(* IEC 61131-3 sources: Elmo_Master/Lasal_PRG/Welcon8Axis_EtherCAT_Test_With_RobotAxis/Class/SafetyCDIAS_Base (part 6) *)

  //Check pointer
  if pData then
    //Length of Firmwareversion (HDINT) -> 8Byte +1 byte zero termination
    if Length >= 9 then
      _itoa(udNumber:=FW_Version, pString:=pData);
    else
      pData^ := 0;
    end_if;
  end_if;

END_FUNCTION

FUNCTION VIRTUAL GLOBAL SafetyCDIAS_Base::GetDiagConnect::NewInst
	VAR_INPUT
		pPara 	  : ^CmdStruct;
		pResult 	: ^Results;
	END_VAR
	VAR_OUTPUT
		ret_code 	: IprStates;
	END_VAR

	ret_code := READY;

	CASE pPara^.uiCmd OF

    CMD_SM_DIAG_GET_INFO:

      //Subcommand
      case pPara^.aPara[0] of
//*****************************************************************************
        SBCMD_SM_DIAG_GET_INFO:
          pResult^.aData[0] :=  GetDiagInfo(pDiagInfo:=(pPara^.aPara[1])$^SafetyDiagInfo);

//*****************************************************************************
        SBCMD_SM_DIAG_GET_STATE:
          pResult^.aData[0] :=  GetDiagState(pDiagState:=(pPara^.aPara[1])$^SafetyDiagState);

//*****************************************************************************
        SBCMD_SM_DIAG_FETCH_INFO:
          //Fetch Diag Info for uCx
          FetchDiagInfo(ucChoice:=pPara^.aPara[1]$USINT);

//*****************************************************************************
        SBCMD_SM_DIAG_FETCH_STATE:
          FetchDiagState();

//*****************************************************************************
        SBCMD_SM_DIAG_IS_SAVE_LOG_ACTIVE:
          pResult^.aData[0] := SaveLogActive();

//*****************************************************************************
        SBCMD_SM_DIAG_SAVE_LOGFILE:
          pResult^.aData[0] := (SaveLog(ucChoice:=(pPara^.aPara[1])$USINT, pDPNE:=(pPara^.aPara[2])$^CHAR))$USINT;

//*****************************************************************************
        SBCMD_SM_DIAG_GET_SAVE_LOGFILE_STATE:
          pResult^.aData[0] := DiagVars.SavingLogSuccessful$USINT;

//*****************************************************************************
        SBCMD_SM_DIAG_GET_SAFETY_NUMBER:
          pResult^.aData[0]$UDINT := SafetyNumber;

//*****************************************************************************
        SBCMD_SM_DIAG_GET_SAFETY_STATE:
          pResult^.aData[0] := ClassState$USINT;

//*****************************************************************************
        SBCMD_SM_DIAG_IS_DIAGNOSE_AVAILABLE:
          pResult^.aData[0] := TRUE;

//*****************************************************************************
        SBCMD_SM_DIAG_GET_CHANNEL_INFO:
          pResult^.aData[0] := GetChannelInfo(pErrorMemUser:=(pPara^.aPara[1])$^UINT, pErrorMem:=#aErrorMem[1], ErrorDataLength:=aErrorMem[0] - 1);
          pResult^.aData[1] := aErrorMem[0] - 1;

//*****************************************************************************
        SBCMD_SM_DIAG_FETCH_CHANNEL_INFO:
          FetchChannelInfo();

//*****************************************************************************
        SBCMD_SM_DIAG_GET_ERRORCODE_OFFSET:

          //Check for valid version
          if pPara^.aPara[1] = 0x01 then  //Version

            ret_code := READY;
            pResult^.aData[0] := 0x01;  //return version
            pResult^.aData[1]$UDINT := GetDiagVisualOffsetErrorCode();

            pResult^.uiLng := 12;

          else

            //invalid version, return error
            ret_code := 1$IprStates; //means iprStates::ERROR but a server error also exists

            pResult^.aData[0] := 0x0;
            pResult^.uiLng    := 4;

          end_if;

      end_case;
    else
      TRACE("(SafetyCDIAS_Base::GetDiagConnect::NewInst) Unknown command!");
      ret_code := 1$IprStates; //means iprStates::ERROR but a server error also exists

	END_CASE;

END_FUNCTION

FUNCTION VIRTUAL GLOBAL SafetyCDIAS_Base::FetchChannelInfo

  DiagVars.UserErrorInfoReady := FALSE;
  DiagVars.UserWantsErrorInfo := TRUE;

END_FUNCTION

FUNCTION VIRTUAL SafetyCDIAS_Base::GetChannelInfo
	VAR_INPUT
		pErrorMemUser 	: ^UINT;
		pErrorMem 	: ^USINT;
		ErrorDataLength 	: INT;
	END_VAR
	VAR_OUTPUT
		StateReady 	: BOOL;
	END_VAR
  VAR
	i   : INT;
  END_VAR

  StateReady := DiagVars.UserErrorInfoReady;

  if StateReady then
    //copy error values in UserArray
    for i := 0 to ErrorDataLength-1 do

      pErrorMemUser^ := pErrorMem^;

      //set pointer to next entry
      pErrorMemUser += sizeof(UINT);
      pErrorMem += sizeof(USINT);
    end_for;
  end_if;

END_FUNCTION

FUNCTION VIRTUAL SafetyCDIAS_Base::GetDiagVisualOffsetErrorCode
	VAR_OUTPUT
		udOffset 	: UDINT;
	END_VAR

  //In the safety firmware for the CSCP and SCP there is only one byte for the errorcode
  //To have different errorcodes (between CSCP and SCP) the safetydesigner adds a fix offset of 1000 to the errorcodes of the SCP01x and SCP11x
  udOffset := 0;

END_FUNCTION
